// TIA Portal V19 export
TYPE "PidL.Feature"
   STRUCT
      Startup : Bool := TRUE;
      MSSOff : Bool := TRUE;
      FltOff : Bool := TRUE;
      LocalMod : Bool;   // 0=Local with Inputs; 1=Local with Feedback
   END_STRUCT;
END_TYPE
